TYPE "ST_PressDemoSignals"
VERSION : 0.1
   STRUCT
      "PartQuality" {ExternalAccessible := 'False'; ExternalVisible := 'False'; ExternalWritable := 'False'} : Bool;
      "AirPressureOk" {ExternalAccessible := 'False'; ExternalVisible := 'False'; ExternalWritable := 'False'} : Bool;
      "PermitDiagnostic" {ExternalAccessible := 'False'; ExternalVisible := 'False'; ExternalWritable := 'False'} : "ST_Diagnostic";
   END_STRUCT;
END_TYPE
